(* LS Electric XG5000 project: NewProject *)
(* PLC LSPLC *)

FUNCTION UserDouble : DINT
(* Doubles an integer *)
VAR_INPUT
    Value : DINT;
END_VAR
UserDouble := Value * 2;
END_FUNCTION

FUNCTION_BLOCK UserAccumulator
(* State retained by each instance between calls *)
VAR_INPUT
    Reset : BOOL;
    Increment : DINT;
END_VAR
VAR_OUTPUT
    Total : DINT;
END_VAR
IF Reset THEN
    Total := 0;
ELSE
    Total := Total + Increment;
END_IF;
END_FUNCTION_BLOCK

PROGRAM NewProgram (* task: 스캔 프로그램 *)
VAR
    Counter : UserAccumulator;
    Observed : DINT;
    Result : DINT;
END_VAR
Result := UserDouble(Value := 4);
Counter(Reset := FALSE, Increment := Result);
Observed := Counter.Total;
END_PROGRAM